// TIA Portal V19 export
DATA_BLOCK "PID_PARAMETERS"   // DB88
{ S7_Optimized_Access := 'FALSE' }
   VAR RETAIN
      R1 : "PID";
      R2 { S7_SetPoint := 'True'} : "PID";
      R3 { S7_SetPoint := 'True'} : "PID";
      R4 { S7_SetPoint := 'True'} : "PID";
      R5 { S7_SetPoint := 'True'} : "PID";
      R6 { S7_SetPoint := 'True'} : "PID";
      R7 { S7_SetPoint := 'True'} : "PID";
      R8 { S7_SetPoint := 'True'} : "PID";
      R9 { S7_SetPoint := 'True'} : "PID";
      R10 { S7_SetPoint := 'True'} : "PID";
      R11 { S7_SetPoint := 'True'} : "PID";
      R12 { S7_SetPoint := 'True'} : "PID";
      R13 { S7_SetPoint := 'True'} : "PID";
      R14 { S7_SetPoint := 'True'} : "PID";
      R15 { S7_SetPoint := 'True'} : "PID";
      R16 { S7_SetPoint := 'True'} : "PID";
      R17 { S7_SetPoint := 'True'} : "PID";
      R18 { S7_SetPoint := 'True'} : "PID";
      HOT_SKID_CP01 { S7_SetPoint := 'True'} : "PID";
      HOT_SKID_CP02 { S7_SetPoint := 'True'} : "PID";
      HOT_SKID_CP03 { S7_SetPoint := 'True'} : "PID";
      COLD_SKID_CP01 { S7_SetPoint := 'True'} : "PID";
      COLD_SKID_CP02 { S7_SetPoint := 'True'} : "PID";
      COLD_SKID_CP03 { S7_SetPoint := 'True'} : "PID";
      CHILLED_SKID_CP01 { S7_SetPoint := 'True'} : "PID";
      CHILLED_SKID_CP02 { S7_SetPoint := 'True'} : "PID";
      CHILLED_SKID_CP03 { S7_SetPoint := 'True'} : "PID";
      ULTRA_CHILLED_SKID_CP01 { S7_SetPoint := 'True'} : "PID";
      ULTRA_CHILLED_SKID_CP02 { S7_SetPoint := 'True'} : "PID";
      HOT_SKID_CV { S7_SetPoint := 'True'} : "PID";
   END_VAR
BEGIN
   R1.P := 0.5;
   R1.I := 1.5;
   R2.P := 0.5;
   R2.I := 1.5;
   R3.P := 0.5;
   R3.I := 1.5;
   R4.P := 0.5;
   R4.I := 1.5;
   R5.P := 0.5;
   R5.I := 1.5;
   R6.P := 0.5;
   R6.I := 1.5;
   R7.P := 0.5;
   R7.I := 1.5;
   R8.P := 0.5;
   R8.I := 1.5;
   R9.P := 0.5;
   R9.I := 1.5;
   R10.P := 0.5;
   R10.I := 1.5;
   R11.P := 0.5;
   R11.I := 1.5;
   R12.P := 0.5;
   R12.I := 1.5;
   R13.P := 0.5;
   R13.I := 1.5;
   R14.P := 0.5;
   R14.I := 1.5;
   R15.P := 0.5;
   R15.I := 1.5;
   R16.P := 0.5;
   R16.I := 1.5;
   R17.P := 0.5;
   R17.I := 1.5;
   R18.P := 0.5;
   R18.I := 1.5;
   HOT_SKID_CP01.P := 0.5;
   HOT_SKID_CP01.I := 1.5;
   HOT_SKID_CP02.P := 0.5;
   HOT_SKID_CP02.I := 1.5;
   HOT_SKID_CP03.P := 0.5;
   HOT_SKID_CP03.I := 1.5;
   COLD_SKID_CP01.P := 0.5;
   COLD_SKID_CP01.I := 1.5;
   COLD_SKID_CP02.P := 0.5;
   COLD_SKID_CP02.I := 1.5;
   COLD_SKID_CP03.P := 0.5;
   COLD_SKID_CP03.I := 1.5;
   CHILLED_SKID_CP01.P := 0.5;
   CHILLED_SKID_CP01.I := 1.5;
   CHILLED_SKID_CP02.P := 0.5;
   CHILLED_SKID_CP02.I := 1.5;
   CHILLED_SKID_CP03.P := 0.5;
   CHILLED_SKID_CP03.I := 1.5;
   ULTRA_CHILLED_SKID_CP01.P := 0.5;
   ULTRA_CHILLED_SKID_CP01.I := 1.5;
   ULTRA_CHILLED_SKID_CP02.P := 0.5;
   ULTRA_CHILLED_SKID_CP02.I := 1.5;
   HOT_SKID_CV.P := 0.5;
   HOT_SKID_CV.I := 1.5;
END_DATA_BLOCK
